Staubli VAL3: actionData.dtx

public actItem aActItem[20]
  [0]
    actionItem aActItem[6]
      [0]
        bool bActive
        num nIOindex = -1
        num nPulseValue
        num nboolValue
        string sIOtype
        string sValue
      [1]
        bool bActive
        num nIOindex = -1
        num nPulseValue
        num nboolValue
        string sIOtype
        string sValue
      [2]
        bool bActive
        num nIOindex = -1
        num nPulseValue
        num nboolValue
        string sIOtype
        string sValue
      [3]
        bool bActive
        num nIOindex = -1
        num nPulseValue
        num nboolValue
        string sIOtype
        string sValue
      [4]
        bool bActive
        num nIOindex = -1
        num nPulseValue
        num nboolValue
        string sIOtype
        string sValue
      [5]
        bool bActive
        num nIOindex = -1
        num nPulseValue
        num nboolValue
        string sIOtype
        string sValue
    string sComment
  [1]
    actionItem aActItem[6]
      [0]
        bool bActive = true
        num nIOindex = 42
        num nPulseValue
        num nboolValue
        string sIOtype = "OUT"
        string sValue = "OFF"
      [1]
        bool bActive = true
        num nIOindex = 43
        num nPulseValue
        num nboolValue
        string sIOtype = "OUT"
        string sValue = "OFF"
      [2]
        bool bActive = true
        num nIOindex = 40
        num nPulseValue
        num nboolValue
        string sIOtype = "OUT"
        string sValue = "OFF"
      [3]
        bool bActive
        num nIOindex = -1
        num nPulseValue
        num nboolValue
        string sIOtype = "OUT"
        string sValue = "ON"
      [4]
        bool bActive
        num nIOindex = -1
        num nPulseValue
        num nboolValue
        string sIOtype = "OUT"
        string sValue = "ON"
      [5]
        bool bActive
        num nIOindex = -1
        num nPulseValue
        num nboolValue
        string sIOtype = "OUT"
        string sValue = "ON"
    string sComment = "int"
  [2]
    actionItem aActItem[6]
      [0]
        bool bActive
        num nIOindex = -1
        num nPulseValue = 0.5
        num nboolValue
        string sIOtype = "PULSE"
        string sValue = "ON"
      [1]
        bool bActive
        num nIOindex = -1
        num nPulseValue
        num nboolValue
        string sIOtype = "OUT"
        string sValue = "OFF"
      [2]
        bool bActive
        num nIOindex = -1
        num nPulseValue
        num nboolValue
        string sIOtype
        string sValue
      [3]
        bool bActive
        num nIOindex = -1
        num nPulseValue
        num nboolValue
        string sIOtype
        string sValue
      [4]
        bool bActive
        num nIOindex = -1
        num nPulseValue
        num nboolValue
        string sIOtype
        string sValue
      [5]
        bool bActive
        num nIOindex = -1
        num nPulseValue
        num nboolValue
        string sIOtype
        string sValue
    string sComment = "action2"
  [3]
    actionItem aActItem[6]
      [0]
        bool bActive
        num nIOindex = -1
        num nPulseValue
        num nboolValue
        string sIOtype
        string sValue
      [1]
        bool bActive
        num nIOindex = -1
        num nPulseValue
        num nboolValue
        string sIOtype
        string sValue
      [2]
        bool bActive
        num nIOindex = -1
        num nPulseValue
        num nboolValue
        string sIOtype
        string sValue
      [3]
        bool bActive
        num nIOindex = -1
        num nPulseValue
        num nboolValue
        string sIOtype
        string sValue
      [4]
        bool bActive
        num nIOindex = -1
        num nPulseValue
        num nboolValue
        string sIOtype
        string sValue
      [5]
        bool bActive
        num nIOindex = -1
        num nPulseValue
        num nboolValue
        string sIOtype
        string sValue
    string sComment = "Action3"
  [4]
    actionItem aActItem[6]
      [0]
        bool bActive
        num nIOindex = -1
        num nPulseValue
        num nboolValue
        string sIOtype
        string sValue
      [1]
        bool bActive
        num nIOindex = -1
        num nPulseValue
        num nboolValue
        string sIOtype
        string sValue
      [2]
        bool bActive
        num nIOindex = -1
        num nPulseValue
        num nboolValue
        string sIOtype
        string sValue
      [3]
        bool bActive
        num nIOindex = -1
        num nPulseValue
        num nboolValue
        string sIOtype
        string sValue
      [4]
        bool bActive
        num nIOindex = -1
        num nPulseValue
        num nboolValue
        string sIOtype
        string sValue
      [5]
        bool bActive
        num nIOindex = -1
        num nPulseValue
        num nboolValue
        string sIOtype
        string sValue
    string sComment = "Action4"
  [5]
    actionItem aActItem[6]
      [0]
        bool bActive
        num nIOindex = -1
        num nPulseValue
        num nboolValue
        string sIOtype
        string sValue
      [1]
        bool bActive
        num nIOindex = -1
        num nPulseValue
        num nboolValue
        string sIOtype
        string sValue
      [2]
        bool bActive
        num nIOindex = -1
        num nPulseValue
        num nboolValue
        string sIOtype
        string sValue
      [3]
        bool bActive
        num nIOindex = -1
        num nPulseValue
        num nboolValue
        string sIOtype
        string sValue
      [4]
        bool bActive
        num nIOindex = -1
        num nPulseValue
        num nboolValue
        string sIOtype
        string sValue
      [5]
        bool bActive
        num nIOindex = -1
        num nPulseValue
        num nboolValue
        string sIOtype
        string sValue
    string sComment = "Action5"
  [6]
    actionItem aActItem[6]
      [0]
        bool bActive
        num nIOindex = -1
        num nPulseValue
        num nboolValue
        string sIOtype
        string sValue
      [1]
        bool bActive
        num nIOindex = -1
        num nPulseValue
        num nboolValue
        string sIOtype
        string sValue
      [2]
        bool bActive
        num nIOindex = -1
        num nPulseValue
        num nboolValue
        string sIOtype
        string sValue
      [3]
        bool bActive
        num nIOindex = -1
        num nPulseValue
        num nboolValue
        string sIOtype
        string sValue
      [4]
        bool bActive
        num nIOindex = -1
        num nPulseValue
        num nboolValue
        string sIOtype
        string sValue
      [5]
        bool bActive
        num nIOindex = -1
        num nPulseValue
        num nboolValue
        string sIOtype
        string sValue
    string sComment = "Action6"
  [7]
    actionItem aActItem[6]
      [0]
        bool bActive
        num nIOindex = -1
        num nPulseValue
        num nboolValue
        string sIOtype
        string sValue
      [1]
        bool bActive
        num nIOindex = -1
        num nPulseValue
        num nboolValue
        string sIOtype
        string sValue
      [2]
        bool bActive
        num nIOindex = -1
        num nPulseValue
        num nboolValue
        string sIOtype
        string sValue
      [3]
        bool bActive
        num nIOindex = -1
        num nPulseValue
        num nboolValue
        string sIOtype
        string sValue
      [4]
        bool bActive
        num nIOindex = -1
        num nPulseValue
        num nboolValue
        string sIOtype
        string sValue
      [5]
        bool bActive
        num nIOindex = -1
        num nPulseValue
        num nboolValue
        string sIOtype
        string sValue
    string sComment = "Action7"
  [8]
    actionItem aActItem[6]
      [0]
        bool bActive
        num nIOindex = -1
        num nPulseValue
        num nboolValue
        string sIOtype
        string sValue
      [1]
        bool bActive
        num nIOindex = -1
        num nPulseValue
        num nboolValue
        string sIOtype
        string sValue
      [2]
        bool bActive
        num nIOindex = -1
        num nPulseValue
        num nboolValue
        string sIOtype
        string sValue
      [3]
        bool bActive
        num nIOindex = -1
        num nPulseValue
        num nboolValue
        string sIOtype
        string sValue
      [4]
        bool bActive
        num nIOindex = -1
        num nPulseValue
        num nboolValue
        string sIOtype
        string sValue
      [5]
        bool bActive
        num nIOindex = -1
        num nPulseValue
        num nboolValue
        string sIOtype
        string sValue
    string sComment = "Action8"
  [9]
    actionItem aActItem[6]
      [0]
        bool bActive
        num nIOindex = -1
        num nPulseValue
        num nboolValue
        string sIOtype
        string sValue
      [1]
        bool bActive
        num nIOindex = -1
        num nPulseValue
        num nboolValue
        string sIOtype
        string sValue
      [2]
        bool bActive
        num nIOindex = -1
        num nPulseValue
        num nboolValue
        string sIOtype
        string sValue
      [3]
        bool bActive
        num nIOindex = -1
        num nPulseValue
        num nboolValue
        string sIOtype
        string sValue
      [4]
        bool bActive
        num nIOindex = -1
        num nPulseValue
        num nboolValue
        string sIOtype
        string sValue
      [5]
        bool bActive
        num nIOindex = -1
        num nPulseValue
        num nboolValue
        string sIOtype
        string sValue
    string sComment = "Action9"
  [10]
    actionItem aActItem[6]
      [0]
        bool bActive
        num nIOindex = -1
        num nPulseValue
        num nboolValue
        string sIOtype
        string sValue
      [1]
        bool bActive
        num nIOindex = -1
        num nPulseValue
        num nboolValue
        string sIOtype
        string sValue
      [2]
        bool bActive
        num nIOindex = -1
        num nPulseValue
        num nboolValue
        string sIOtype
        string sValue
      [3]
        bool bActive
        num nIOindex = -1
        num nPulseValue
        num nboolValue
        string sIOtype
        string sValue
      [4]
        bool bActive
        num nIOindex = -1
        num nPulseValue
        num nboolValue
        string sIOtype
        string sValue
      [5]
        bool bActive
        num nIOindex = -1
        num nPulseValue
        num nboolValue
        string sIOtype
        string sValue
    string sComment = "Action10"
  [11]
    actionItem aActItem[6]
      [0]
        bool bActive
        num nIOindex = -1
        num nPulseValue
        num nboolValue
        string sIOtype
        string sValue
      [1]
        bool bActive
        num nIOindex = -1
        num nPulseValue
        num nboolValue
        string sIOtype
        string sValue
      [2]
        bool bActive
        num nIOindex = -1
        num nPulseValue
        num nboolValue
        string sIOtype
        string sValue
      [3]
        bool bActive
        num nIOindex = -1
        num nPulseValue
        num nboolValue
        string sIOtype
        string sValue
      [4]
        bool bActive
        num nIOindex = -1
        num nPulseValue
        num nboolValue
        string sIOtype
        string sValue
      [5]
        bool bActive
        num nIOindex = -1
        num nPulseValue
        num nboolValue
        string sIOtype
        string sValue
    string sComment = "Action11"
  [12]
    actionItem aActItem[6]
      [0]
        bool bActive
        num nIOindex = -1
        num nPulseValue
        num nboolValue
        string sIOtype
        string sValue
      [1]
        bool bActive
        num nIOindex = -1
        num nPulseValue
        num nboolValue
        string sIOtype
        string sValue
      [2]
        bool bActive
        num nIOindex = -1
        num nPulseValue
        num nboolValue
        string sIOtype
        string sValue
      [3]
        bool bActive
        num nIOindex = -1
        num nPulseValue
        num nboolValue
        string sIOtype
        string sValue
      [4]
        bool bActive
        num nIOindex = -1
        num nPulseValue
        num nboolValue
        string sIOtype
        string sValue
      [5]
        bool bActive
        num nIOindex = -1
        num nPulseValue
        num nboolValue
        string sIOtype
        string sValue
    string sComment = "Action12"
  [13]
    actionItem aActItem[6]
      [0]
        bool bActive
        num nIOindex = -1
        num nPulseValue
        num nboolValue
        string sIOtype
        string sValue
      [1]
        bool bActive
        num nIOindex = -1
        num nPulseValue
        num nboolValue
        string sIOtype
        string sValue
      [2]
        bool bActive
        num nIOindex = -1
        num nPulseValue
        num nboolValue
        string sIOtype
        string sValue
      [3]
        bool bActive
        num nIOindex = -1
        num nPulseValue
        num nboolValue
        string sIOtype
        string sValue
      [4]
        bool bActive
        num nIOindex = -1
        num nPulseValue
        num nboolValue
        string sIOtype
        string sValue
      [5]
        bool bActive
        num nIOindex = -1
        num nPulseValue
        num nboolValue
        string sIOtype
        string sValue
    string sComment = "Action13"
  [14]
    actionItem aActItem[6]
      [0]
        bool bActive
        num nIOindex = -1
        num nPulseValue
        num nboolValue
        string sIOtype
        string sValue
      [1]
        bool bActive
        num nIOindex = -1
        num nPulseValue
        num nboolValue
        string sIOtype
        string sValue
      [2]
        bool bActive
        num nIOindex = -1
        num nPulseValue
        num nboolValue
        string sIOtype
        string sValue
      [3]
        bool bActive
        num nIOindex = -1
        num nPulseValue
        num nboolValue
        string sIOtype
        string sValue
      [4]
        bool bActive
        num nIOindex = -1
        num nPulseValue
        num nboolValue
        string sIOtype
        string sValue
      [5]
        bool bActive
        num nIOindex = -1
        num nPulseValue
        num nboolValue
        string sIOtype
        string sValue
    string sComment = "Action14"
  [15]
    actionItem aActItem[6]
      [0]
        bool bActive
        num nIOindex = 16
        num nPulseValue
        num nboolValue
        string sIOtype = "OUT"
        string sValue = "ON"
      [1]
        bool bActive
        num nIOindex = 18
        num nPulseValue
        num nboolValue
        string sIOtype = "OUT"
        string sValue = "OFF"
      [2]
        bool bActive
        num nIOindex = -1
        num nPulseValue
        num nboolValue
        string sIOtype
        string sValue
      [3]
        bool bActive
        num nIOindex = -1
        num nPulseValue
        num nboolValue
        string sIOtype
        string sValue
      [4]
        bool bActive
        num nIOindex = -1
        num nPulseValue
        num nboolValue
        string sIOtype
        string sValue
      [5]
        bool bActive
        num nIOindex = -1
        num nPulseValue
        num nboolValue
        string sIOtype
        string sValue
    string sComment = "Action15"
  [16]
    actionItem aActItem[6]
      [0]
        bool bActive
        num nIOindex = -1
        num nPulseValue
        num nboolValue
        string sIOtype
        string sValue
      [1]
        bool bActive
        num nIOindex = -1
        num nPulseValue
        num nboolValue
        string sIOtype
        string sValue
      [2]
        bool bActive
        num nIOindex = -1
        num nPulseValue
        num nboolValue
        string sIOtype
        string sValue
      [3]
        bool bActive
        num nIOindex = -1
        num nPulseValue
        num nboolValue
        string sIOtype
        string sValue
      [4]
        bool bActive
        num nIOindex = -1
        num nPulseValue
        num nboolValue
        string sIOtype
        string sValue
      [5]
        bool bActive
        num nIOindex = -1
        num nPulseValue
        num nboolValue
        string sIOtype
        string sValue
    string sComment = "Action16"
  [17]
    actionItem aActItem[6]
      [0]
        bool bActive
        num nIOindex = -1
        num nPulseValue
        num nboolValue
        string sIOtype
        string sValue
      [1]
        bool bActive
        num nIOindex = -1
        num nPulseValue
        num nboolValue
        string sIOtype
        string sValue
      [2]
        bool bActive
        num nIOindex = -1
        num nPulseValue
        num nboolValue
        string sIOtype
        string sValue
      [3]
        bool bActive
        num nIOindex = -1
        num nPulseValue
        num nboolValue
        string sIOtype
        string sValue
      [4]
        bool bActive
        num nIOindex = -1
        num nPulseValue
        num nboolValue
        string sIOtype
        string sValue
      [5]
        bool bActive
        num nIOindex = -1
        num nPulseValue
        num nboolValue
        string sIOtype
        string sValue
    string sComment = "Action17"
  [18]
    actionItem aActItem[6]
      [0]
        bool bActive
        num nIOindex = -1
        num nPulseValue
        num nboolValue
        string sIOtype
        string sValue
      [1]
        bool bActive
        num nIOindex = -1
        num nPulseValue
        num nboolValue
        string sIOtype
        string sValue
      [2]
        bool bActive
        num nIOindex = -1
        num nPulseValue
        num nboolValue
        string sIOtype
        string sValue
      [3]
        bool bActive
        num nIOindex = -1
        num nPulseValue
        num nboolValue
        string sIOtype
        string sValue
      [4]
        bool bActive
        num nIOindex = -1
        num nPulseValue
        num nboolValue
        string sIOtype
        string sValue
      [5]
        bool bActive
        num nIOindex = -1
        num nPulseValue
        num nboolValue
        string sIOtype
        string sValue
    string sComment = "Action18"
  [19]
    actionItem aActItem[6]
      [0]
        bool bActive
        num nIOindex = -1
        num nPulseValue
        num nboolValue
        string sIOtype
        string sValue
      [1]
        bool bActive
        num nIOindex = -1
        num nPulseValue
        num nboolValue
        string sIOtype
        string sValue
      [2]
        bool bActive
        num nIOindex = -1
        num nPulseValue
        num nboolValue
        string sIOtype
        string sValue
      [3]
        bool bActive
        num nIOindex = -1
        num nPulseValue
        num nboolValue
        string sIOtype
        string sValue
      [4]
        bool bActive
        num nIOindex = -1
        num nPulseValue
        num nboolValue
        string sIOtype
        string sValue
      [5]
        bool bActive
        num nIOindex = -1
        num nPulseValue
        num nboolValue
        string sIOtype
        string sValue
    string sComment = "Action19"
